FUNCTION_BLOCK FB_EL3351Measuring_1
VAR_INPUT
(*+++++ Inputs from Device +++++*)
	diDiffvoltage: DINT;
	diRefvoltage: DINT;

END_VAR
VAR_OUTPUT
	rUref: REAL;
	rUdiff: REAL;
	rGrossWeight: REAL;
	rNetWeight: REAL;
	rTareWeight: REAL;
END_VAR
VAR
(*+++++ Inputs that can be made in the visu +++++*)
	rRatedOutput: REAL;
	rRatedCapacity: REAL;
	rZeroBalance: REAL;
(*+++++ Values that are needed to do calculations  +++++*)
	rRefvoltageConv: REAL;
	rDiffvoltageConv: REAL;
(*+++++ Visu Buttons / Strings +++++*)
	fbRTrig_SetTare: R_TRIG;
	fbRTrig_ResetTare: R_TRIG;
	bSetTare: BOOL;
	bResetTare: BOOL;
	sSettings: STRING(150);
(*+++++ Auto Calibration +++++*)
	bCalibration: BOOL;
	bStartCalibration: BOOL;
	fbRTrig_StartCalibration: R_TRIG;
	bNextStep: BOOL;
	fbRTrig_NextStep: R_TRIG;
	nStepCalibrate: UDINT;
	rReferenceWeight: REAL;
	rOffset: REAL;
	rCalculatedRatedOutput: REAL;
	rUdiffWithoutOffset: REAL;
	sRatedCapacity: STRING;
END_VAR
VAR CONSTANT
	rVoltageSupply				:REAL := 12.0;			(* [V] *)
	rSensorType					:REAL := 20.0;			(* [mV] *)
END_VAR


(*For being able to do calculations, the Inputs from the device need to be converted to REAL values*)
rRefvoltageConv:= DINT_TO_REAL(diRefvoltage);
rDiffvoltageConv:= DINT_TO_REAL(diDiffvoltage);

(*Calculation of Voltages*)
rUref:= rRefvoltageConv*(rVoltageSupply/2147483647);
rUdiff:= rDiffvoltageConv*(rSensorType/2147483647);

(*++++++++++++++++++++++++++++++ Manual Mode +++++++++++++++++++++++++++++*)
IF NOT bCalibration THEN									(*Settings can be changed manually by default*)
	nStepCalibrate:= 0;
	sSettings:= 'Settings can be changed manually! ';
	IF rRatedCapacity= 0												(*It is checked if inputs have yet been made*)
	THEN
		sSettings:=  CONCAT(sSettings, 'Enter Rated Capacity! ');
	END_IF

	IF rRatedOutput = 0 THEN
		sSettings:= CONCAT(sSettings, 'Enter Rated Output! ');
	END_IF
	sSettings:= CONCAT(sSettings, '$n');
	sSettings:= CONCAT(sSettings, 'If you want Settings to be set automatically, activate Calibration Mode. ');
END_IF

(*++++++++++++++++++++++++++++++ Calibration Mode +++++++++++++++++++++++++++++*)
IF bCalibration THEN
	CASE nStepCalibrate OF

		0:	(*Calibration is started, when button "Start Calibration" is pressed. As long as it hasn't been pressed, the button blinks blue *)
			IF NOT fbRTrig_StartCalibration.Q THEN
				sSettings:= 'Calibration Mode ON. Press Start Calibration or deactivate Calibration Mode. ';
			ELSE
				nStepCalibrate:= nStepCalibrate+10;
			END_IF
	
		10:	(*First of all it is checked, if the Rated Capacity has yet been typed in. If not, the shape blinks blue.
			If some value has been typed in, the user is asked, whether it is correct. Pressing "Save" starts the next step. *)
			rGrossWeight:= 0;
			rOffset:= 0;
			rCalculatedRatedOutput:= 0;
			rReferenceWeight:= 0;
			IF rRatedCapacity= 0 THEN
				sSettings:= 'Calibration Mode ON. Enter Rated Capacity of Load Cell! Then press Save! ';
			ELSIF rRatedCapacity <> 0 THEN
				sSettings:= 'Calibration Mode ON. If Rated Capacity of ';
				sRatedCapacity:= REAL_TO_STRING(rRatedCapacity);
				sSettings:= CONCAT(sSettings, sRatedCapacity);
				sSettings:= CONCAT(sSettings, 'kg is correct, press Save! ');
				IF fbRTrig_NextStep.Q THEN
					nStepCalibrate:= nStepCalibrate+10;
				END_IF
			END_IF
	
		20:	(*The Zero Balance of the load cell is detected. Therefore, no load must be put on the load cell. *)
			sSettings:= 'Remove all load from load cell! Then press Save! ';
			IF fbRTrig_NextStep.Q THEN
				rOffset:= rUdiff/rUref;
				rZeroBalance:= rOffset;
				nStepCalibrate:= nStepCalibrate+10;
			END_IF

			IF fbRTrig_StartCalibration.Q THEN
				nStepCalibrate:= 10;
			END_IF
	
		30:	(*The Rated Output is detected. Therefore, a reference weight must be put on the load cell and it must be entered.*)
			sSettings:= 'Put Reference Weight on load cell! Enter reference weight! Then press Save! ';
			IF rReferenceWeight <> 0 THEN
				sSettings:= 'Make sure reference weight is on load cell! Then press Save! ';
				IF fbRTrig_NextStep.Q THEN
					rCalculatedRatedOutput:= (rUdiffWithoutOffset/rUref)*(rRatedCapacity/rReferenceWeight);
					rRatedOutput:= rCalculatedRatedOutput;
					nStepCalibrate:= nStepCalibrate+ 10;
				END_IF
			END_IF

			IF fbRTrig_StartCalibration.Q THEN
				nStepCalibrate:= 10;
			END_IF
	
		40:	(*Once the zero balance and the Rated Output have been detected, "Start Calibration" can be pressed to restart the Calibration process*)
			sSettings:= 'Auto Calibration complete. If necessary, press Start Calibration to reconfigure.';
			IF fbRTrig_StartCalibration.Q THEN
				nStepCalibrate:= 10;
			END_IF
			IF rRatedCapacity= 0 THEN
			sSettings:=  CONCAT(sSettings, '$n');
			sSettings:=  CONCAT(sSettings, 'Enter Rated Capacity! ');
			END_IF
	END_CASE
END_IF

(*++++++++++++++++++++++++++++++ Calculation of Weight +++++++++++++++++++++++++++++*)
rUdiffWithoutOffset:= rUdiff-(rZeroBalance*rUref);

IF rRatedOutput<>0 THEN
	rGrossWeight:= (rUdiffWithoutOffset/rUref)*(rRatedCapacity/rRatedOutput);
ELSE
	rGrossWeight:= 0;
END_IF

(*++++++++++++++++++++++++++++++ Tare Weight +++++++++++++++++++++++++++++*)
IF rRatedCapacity <> 0 AND rRatedOutput <> 0 THEN
	fbRTrig_SetTare( CLK:= bSetTare, Q=> );
	IF fbRTrig_SetTare.Q THEN
		rTareWeight:= rGrossWeight;
	END_IF

	IF rTareWeight= 0 THEN
		rNetWeight:= 0;
	ELSE
		rNetWeight:= rGrossWeight- rTareWeight;		(*Calculation of the shown Net Weight*)
	END_IF
END_IF

(*When the Button 'Reset Tare Weight' is pressed, the Tare Value is reset*)
fbRTrig_ResetTare( CLK:= bResetTare, Q=> );
IF fbRTrig_ResetTare.Q THEN
	rTareWeight:= 0;
END_IF


fbRTrig_StartCalibration( CLK:= bStartCalibration, Q=> );
fbRTrig_NextStep( CLK:= bNextStep, Q=> );

END_FUNCTION_BLOCK

(* stored: Version 1.1.0.1, ProductVersion 3.1.4024.15
   POU FB_EL3351Measuring_1: Id {3428cabf-dfd6-499d-a532-62a682926eef}, SpecialFunc None *)
